// Mitsubishi GX Works2 project: 최종_HMIV2   PLC: Q02/Q02H

PROGRAM MAIN
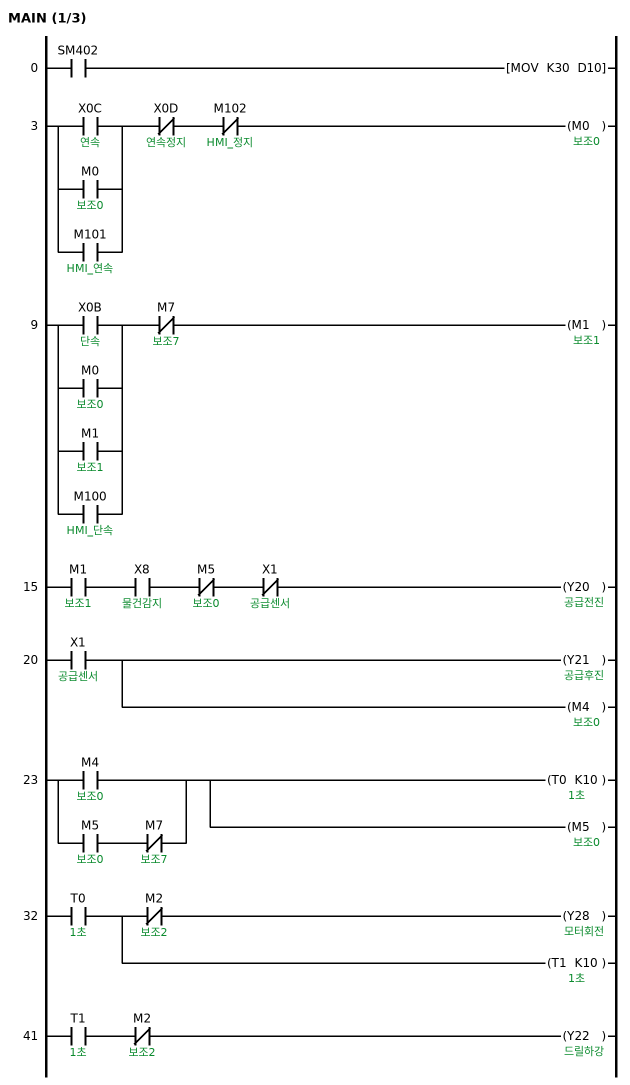
0     LD      SM402
      MOV     K30 D10
3     LD      X0C  ; 연속
      OR      M0  ; 보조0
      OR      M101  ; HMI_연속
      ANI     X0D  ; 연속정지
      ANI     M102  ; HMI_정지
      OUT     M0  ; 보조0
9     LD      X0B  ; 단속
      OR      M0  ; 보조0
      OR      M1  ; 보조1
      OR      M100  ; HMI_단속
      ANI     M7  ; 보조7
      OUT     M1  ; 보조1
15    LD      M1  ; 보조1
      AND     X8  ; 물건감지
      ANI     M5  ; 보조0
      ANI     X1  ; 공급센서
      OUT     Y20  ; 공급전진
20    LD      X1  ; 공급센서
      OUT     Y21  ; 공급후진
      OUT     M4  ; 보조0
23    LD      M4  ; 보조0
      LD      M5  ; 보조0
      ANI     M7  ; 보조7
      ORB
      OUT     T0 K10  ; 1초
      OUT     M5  ; 보조0
32    LD      T0  ; 1초
      MPS
      ANI     M2  ; 보조2
      OUT     Y28  ; 모터회전
      MPP
      OUT     T1 K10  ; 1초
41    LD      T1  ; 1초
      ANI     M2  ; 보조2
      OUT     Y22  ; 드릴하강
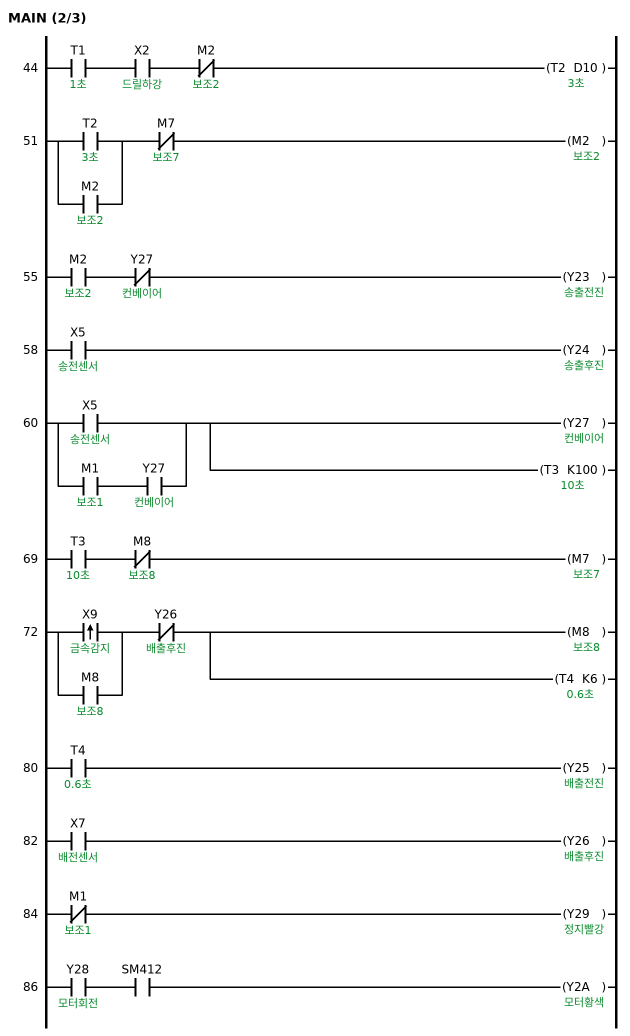
44    LD      T1  ; 1초
      AND     X2  ; 드릴하강
      ANI     M2  ; 보조2
      OUT     T2 D10  ; 3초
51    LD      T2  ; 3초
      OR      M2  ; 보조2
      ANI     M7  ; 보조7
      OUT     M2  ; 보조2
55    LD      M2  ; 보조2
      ANI     Y27  ; 컨베이어
      OUT     Y23  ; 송출전진
58    LD      X5  ; 송전센서
      OUT     Y24  ; 송출후진
60    LD      X5  ; 송전센서
      LD      M1  ; 보조1
      AND     Y27  ; 컨베이어
      ORB
      OUT     Y27  ; 컨베이어
      OUT     T3 K100  ; 10초
69    LD      T3  ; 10초
      ANI     M8  ; 보조8
      OUT     M7  ; 보조7
72    LDP     X9  ; 금속감지
      OR      M8  ; 보조8
      ANI     Y26  ; 배출후진
      OUT     M8  ; 보조8
      OUT     T4 K6  ; 0.6초
80    LD      T4  ; 0.6초
      OUT     Y25  ; 배출전진
82    LD      X7  ; 배전센서
      OUT     Y26  ; 배출후진
84    LDI     M1  ; 보조1
      OUT     Y29  ; 정지빨강
86    LD      Y28  ; 모터회전
      AND     SM412
      OUT     Y2A  ; 모터황색
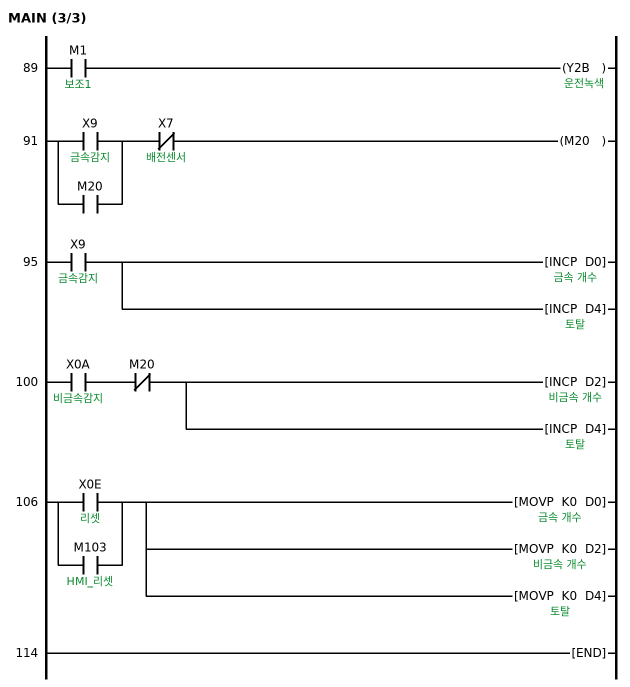
89    LD      M1  ; 보조1
      OUT     Y2B  ; 운전녹색
91    LD      X9  ; 금속감지
      OR      M20
      ANI     X7  ; 배전센서
      OUT     M20
95    LD      X9  ; 금속감지
      INCP    D0  ; 금속 개수
      INCP    D4  ; 토탈
100   LD      X0A  ; 비금속감지
      ANI     M20
      INCP    D2  ; 비금속 개수
      INCP    D4
106   LD      X0E  ; 리셋
      OR      M103  ; HMI_리셋
      MOVP    K0 D0
      MOVP    K0 D2
      MOVP    K0 D4
114   END
END_PROGRAM

PROGRAM LAMP
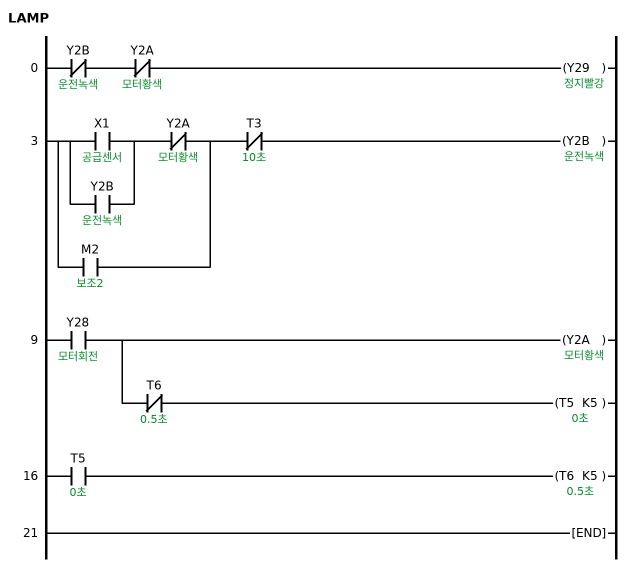
0     LDI     Y2B  ; 운전녹색
      ANI     Y2A  ; 모터황색
      OUT     Y29  ; 정지빨강
3     LD      X1  ; 공급센서
      OR      Y2B  ; 운전녹색
      ANI     Y2A  ; 모터황색
      OR      M2  ; 보조2
      ANI     T3  ; 10초
      OUT     Y2B  ; 운전녹색
9     LD      Y28  ; 모터회전
      OUT     Y2A  ; 모터황색
      ANI     T6  ; 0.5초
      OUT     T5 K5  ; 0초
16    LD      T5  ; 0초
      OUT     T6 K5  ; 0.5초
21    END
END_PROGRAM

// device comments not shown above
X0  ; 공후센서
X6  ; 배후센서
M3  ; 보조3
M6  ; 보조0
M9  ; 보조9
M99  ; 단속정지
